// TIA Portal V19 export
// export: Created 2026-10-15T09:44:24.662474Z, ExportSetting WithDefaults, DisplayName Totally Integrated Automation Portal, DisplayVersion V19, DisplayName TIA Portal Openness, DisplayVersion V19, DisplayName TIA Portal Version Control Interface, DisplayVersion V19, DisplayName STEP 7 Professional, DisplayVersion V19, DisplayName STEP 7 Safety, DisplayVersion V19, DisplayName WinCC Basic/Comfort/Advanced, DisplayVersion V19, DisplayName WinCC Unified, DisplayVersion V19
FUNCTION "ROLL_PB20" : Void   // FC28, SCL
{ S7_Optimized_Access := 'TRUE' }
VERSION : 0.1
// stored: AutoNumber true, IsIECCheckEnabled false, SetENOAutomatically false, UDAEnableTagReadback false
   VAR_TEMP
      r : Bool;
      a1 : Word;
      a2 : Word;
      activeDataBlock : Int;
      comparisonResults : Array[0..0] of Bool;
   END_VAR
BEGIN

   #r := FALSE;
   #a1 := W#16#0000;
   #a2 := W#16#0000;
   #activeDataBlock := 0;
   // PB20, STEP 5 network 1
   #activeDataBlock := 15;
   // PB20, STEP 5 network 2
   #r := ((NOT "ROLL_IO".Input[7, 0]) AND (("ROLL_IO".Input[0, 1] AND "ROLL_State".M[190, 6] AND "ROLL_State".M[26, 5] AND "ROLL_State".M[4, 1]) OR ("ROLL_IO".Input[0, 2] AND "ROLL_State".M[0, 3])) AND "ROLL_State".M[4, 1]);
   "ROLL_State".M[8, 0] := #r;
   // PB20, STEP 5 network 3
   #r := ((NOT "ROLL_IO".Input[7, 1]) AND "ROLL_IO".Input[0, 2] AND "ROLL_IO".Input[1, 6] AND "ROLL_State".M[4, 1] AND "ROLL_State".S5Timers[61].Q);
   IF #r THEN
       "ROLL_State".M[8, 1] := TRUE;
   END_IF;
   #r := "ROLL_State".M[3, 1];
   IF #r THEN
       "ROLL_State".M[8, 1] := FALSE;
   END_IF;
   // PB20, STEP 5 network 4
   #a2 := #a1;
   #a1 := "ROLL_GetDW"(DbNumber := #activeDataBlock, Index := 61);
   #r := ((NOT "ROLL_IO".Input[7, 1]) AND "ROLL_IO".Input[0, 2] AND "ROLL_IO".Input[3, 1]);
   "ROLL_TimerOp"(Number := 61,
                  Operation := 0,
                  Signal := #r,
                  Preset := #a1);
   #r := ("ROLL_State".M[3, 1] AND "ROLL_State".M[4, 1]);
   "ROLL_TimerOp"(Number := 61,
                  Operation := 2,
                  Signal := #r,
                  Preset := #a1);
   // PB20, STEP 5 network 5
   #r := ((NOT "ROLL_IO".Input[7, 2]) AND "ROLL_State".S5Timers[55].Q);
   IF #r THEN
       "ROLL_State".M[8, 2] := TRUE;
   END_IF;
   #r := "ROLL_State".M[3, 1];
   IF #r THEN
       "ROLL_State".M[8, 2] := FALSE;
   END_IF;
   // PB20, STEP 5 network 6
   #a2 := #a1;
   #a1 := "ROLL_GetDW"(DbNumber := #activeDataBlock, Index := 55);
   #r := ((NOT "ROLL_IO".Input[7, 2]) AND (NOT "ROLL_State".M[8, 2]) AND "ROLL_State".M[4, 1]);
   "ROLL_TimerOp"(Number := 55,
                  Operation := 0,
                  Signal := #r,
                  Preset := #a1);
   // PB20, STEP 5 network 7
   #r := ((NOT "ROLL_IO".Input[7, 3]) AND "ROLL_IO".Output[21, 6] AND "ROLL_State".S5Timers[60].Q);
   IF #r THEN
       "ROLL_State".M[8, 3] := TRUE;
   END_IF;
   #r := "ROLL_State".M[3, 1];
   IF #r THEN
       "ROLL_State".M[8, 3] := FALSE;
   END_IF;
   // PB20, STEP 5 network 8
   #a2 := #a1;
   #a1 := "ROLL_GetDW"(DbNumber := #activeDataBlock, Index := 60);
   #r := ((NOT "ROLL_IO".Input[7, 3]) AND "ROLL_IO".Output[21, 6] AND "ROLL_IO".Input[3, 1]);
   "ROLL_TimerOp"(Number := 60,
                  Operation := 0,
                  Signal := #r,
                  Preset := #a1);
   // PB20, STEP 5 network 9
   #a2 := #a1;
   #a1 := W#16#2010;
   #r := (NOT "ROLL_IO".Input[7, 4]);
   "ROLL_TimerOp"(Number := 88,
                  Operation := 0,
                  Signal := #r,
                  Preset := #a1);
   // PB20, STEP 5 network 10
   #r := ((NOT "ROLL_IO".Input[7, 4]) AND "ROLL_State".M[4, 1] AND "ROLL_State".S5Timers[88].Q);
   "ROLL_State".M[8, 4] := #r;
   // PB20, STEP 5 network 11
   #r := (("ROLL_State".M[25, 0] OR "ROLL_State".M[25, 1]) AND "ROLL_IO".Input[0, 1] AND "ROLL_State".M[190, 6] AND "ROLL_State".M[4, 1] AND "ROLL_State".S5Timers[96].Q);
   IF #r THEN
       "ROLL_State".M[8, 5] := TRUE;
   END_IF;
   #r := "ROLL_State".M[3, 1];
   IF #r THEN
       "ROLL_State".M[8, 5] := FALSE;
   END_IF;
   // PB20, STEP 5 network 12
   #r := ((NOT "ROLL_IO".Input[9, 0]) AND ("ROLL_IO".Input[1, 6] OR "ROLL_IO".Input[1, 7]) AND "ROLL_IO".Input[9, 6]);
   IF #r THEN
       "ROLL_State".M[12, 4] := TRUE;
   END_IF;
   #r := "ROLL_State".M[3, 1];
   IF #r THEN
       "ROLL_State".M[12, 4] := FALSE;
   END_IF;
   // PB20, STEP 5 network 13
   #r := ((NOT "ROLL_IO".Input[9, 3]) AND ("ROLL_IO".Input[1, 6] OR "ROLL_IO".Input[1, 7]) AND "ROLL_IO".Input[9, 6]);
   IF #r THEN
       "ROLL_State".M[12, 5] := TRUE;
   END_IF;
   #r := "ROLL_State".M[3, 1];
   IF #r THEN
       "ROLL_State".M[12, 5] := FALSE;
   END_IF;
   // PB20, STEP 5 network 14
   #r := ((NOT "ROLL_IO".Input[9, 7]) AND ("ROLL_IO".Input[1, 6] OR "ROLL_IO".Input[1, 7]));
   IF #r THEN
       "ROLL_State".M[12, 6] := TRUE;
   END_IF;
   #r := "ROLL_State".M[3, 1];
   IF #r THEN
       "ROLL_State".M[12, 6] := FALSE;
   END_IF;
   // PB20, STEP 5 network 15
   #r := (NOT "ROLL_IO".Input[9, 6]);
   IF #r THEN
       "ROLL_State".M[12, 7] := TRUE;
   END_IF;
   #r := ("ROLL_IO".Input[9, 6] AND "ROLL_State".M[3, 1]);
   IF #r THEN
       "ROLL_State".M[12, 7] := FALSE;
   END_IF;
   // PB20, STEP 5 network 16
   #a2 := #a1;
   #a1 := "ROLL_GetDW"(DbNumber := #activeDataBlock, Index := 56);
   #r := (NOT "ROLL_IO".Input[7, 1]);
   "ROLL_TimerOp"(Number := 56,
                  Operation := 1,
                  Signal := #r,
                  Preset := #a1);
   // PB20, STEP 5 network 17
   #a2 := #a1;
   #a1 := "ROLL_GetDW"(DbNumber := #activeDataBlock, Index := 65);
   #r := (NOT "ROLL_IO".Input[7, 3]);
   "ROLL_TimerOp"(Number := 65,
                  Operation := 0,
                  Signal := #r,
                  Preset := #a1);
   // PB20, STEP 5 network 18
   #a2 := #a1;
   #a1 := W#16#2020;
   #r := "ROLL_IO".Input[7, 3];
   "ROLL_TimerOp"(Number := 66,
                  Operation := 1,
                  Signal := #r,
                  Preset := #a1);
   // PB20, STEP 5 network 19
   #a2 := #a1;
   #a1 := "ROLL_GetDW"(DbNumber := #activeDataBlock, Index := 67);
   #r := ("ROLL_IO".Input[7, 3] AND "ROLL_State".M[150, 1]);
   "ROLL_TimerOp"(Number := 67,
                  Operation := 0,
                  Signal := #r,
                  Preset := #a1);
   // PB20, STEP 5 network 20
   #a2 := #a1;
   #a1 := W#16#2005;
   #r := (NOT "ROLL_IO".Input[7, 5]);
   "ROLL_TimerOp"(Number := 96,
                  Operation := 0,
                  Signal := #r,
                  Preset := #a1);
   // PB20, STEP 5 network 21
   #a2 := #a1;
   #a1 := W#16#2030;
   #r := "ROLL_IO".Input[7, 5];
   "ROLL_TimerOp"(Number := 97,
                  Operation := 0,
                  Signal := #r,
                  Preset := #a1);
   // PB20, STEP 5 network 22
   #r := (((NOT "ROLL_IO".Output[18, 5]) AND "ROLL_IO".Output[18, 4]) OR ((NOT "ROLL_IO".Output[18, 7]) AND "ROLL_IO".Output[18, 6]));
   "ROLL_State".M[149, 6] := #r;
   // PB20, STEP 5 network 23
   #a2 := #a1;
   #a1 := W#16#1010;
   #r := "ROLL_State".M[148, 4];
   "ROLL_TimerOp"(Number := 89,
                  Operation := 0,
                  Signal := #r,
                  Preset := #a1);
   // PB20, STEP 5 network 24
   #r := "ROLL_State".M[149, 6];
   IF #r THEN
       "ROLL_State".M[148, 4] := TRUE;
   END_IF;
   #r := "ROLL_State".S5Timers[89].Q;
   IF #r THEN
       "ROLL_State".M[148, 4] := FALSE;
   END_IF;
   // PB20, STEP 5 network 25
   #r := ("ROLL_IO".Input[8, 0] AND "ROLL_State".S5Timers[70].Q);
   "ROLL_State".M[147, 0] := #r;
   // PB20, STEP 5 network 26
   #a2 := #a1;
   #a1 := "ROLL_GetDW"(DbNumber := #activeDataBlock, Index := 75);
   #r := (NOT "ROLL_State".M[147, 0]);
   "ROLL_TimerOp"(Number := 75,
                  Operation := 0,
                  Signal := #r,
                  Preset := #a1);
   // PB20, STEP 5 network 27
   #r := "ROLL_State".M[0, 3];
   "ROLL_State".M[147, 1] := #r;
   // PB20, STEP 5 network 28
   #r := ("ROLL_IO".Input[8, 2] AND "ROLL_State".S5Timers[72].Q);
   "ROLL_State".M[147, 2] := #r;
   // PB20, STEP 5 network 29
   #a2 := #a1;
   #a1 := "ROLL_GetDW"(DbNumber := #activeDataBlock, Index := 77);
   #r := (NOT "ROLL_State".M[147, 2]);
   "ROLL_TimerOp"(Number := 77,
                  Operation := 0,
                  Signal := #r,
                  Preset := #a1);
   // PB20, STEP 5 network 30
   #r := "ROLL_State".M[0, 3];
   "ROLL_State".M[149, 0] := #r;
   // PB20, STEP 5 network 31
   #r := ("ROLL_State".M[147, 0] OR "ROLL_State".M[147, 2]);
   "ROLL_State".M[149, 1] := #r;
   // PB20, STEP 5 network 32
   #r := "ROLL_State".M[0, 3];
   "ROLL_State".M[149, 2] := #r;
   // PB20, STEP 5 network 33
   #r := ("ROLL_State".M[147, 0] AND "ROLL_State".M[147, 2]);
   "ROLL_State".M[149, 3] := #r;
   // PB20, STEP 5 network 34
   #r := ((NOT "ROLL_State".M[12, 6]) AND (NOT "ROLL_State".M[12, 7]) AND (NOT "ROLL_State".M[13, 4]) AND (NOT "ROLL_State".M[6, 0]) AND (NOT "ROLL_State".M[6, 2]) AND (NOT "ROLL_State".M[8, 2]) AND ("ROLL_IO".Input[1, 6] OR "ROLL_IO".Input[1, 7]) AND "ROLL_IO".Input[3, 1] AND "ROLL_IO".Input[7, 4] AND "ROLL_IO".Input[9, 6] AND "ROLL_IO".Input[9, 7] AND "ROLL_State".S5Timers[66].Q);
   "ROLL_State".M[150, 2] := #r;
   // PB20, STEP 5 network 35
   #r := ((NOT "ROLL_IO".Input[9, 2]) AND (NOT "ROLL_State".M[12, 4]) AND ("ROLL_IO".Output[18, 4] OR "ROLL_IO".Input[9, 1]) AND ("ROLL_State".M[149, 0] OR "ROLL_State".M[149, 1] OR "ROLL_State".M[149, 2] OR "ROLL_State".M[149, 3]) AND "ROLL_IO".Input[9, 0] AND "ROLL_State".M[150, 2]);
   "ROLL_IO".Output[18, 4] := #r;
   // PB20, STEP 5 network 36
   #r := ((NOT "ROLL_IO".Input[9, 2]) AND (NOT "ROLL_State".M[12, 4]) AND ("ROLL_IO".Output[18, 4] OR "ROLL_IO".Output[18, 5] OR "ROLL_IO".Input[9, 1]) AND ("ROLL_State".M[149, 2] OR "ROLL_State".M[149, 3]) AND "ROLL_IO".Input[9, 0] AND "ROLL_State".M[150, 2]);
   "ROLL_IO".Output[18, 5] := #r;
   // PB20, STEP 5 network 37
   #r := ((NOT "ROLL_IO".Input[9, 5]) AND (NOT "ROLL_State".M[12, 5]) AND ("ROLL_IO".Output[18, 6] OR "ROLL_IO".Input[9, 4]) AND ("ROLL_State".M[149, 1] OR "ROLL_State".M[149, 2] OR "ROLL_State".M[149, 3]) AND "ROLL_IO".Input[9, 3] AND "ROLL_State".M[150, 2]);
   "ROLL_IO".Output[18, 6] := #r;
   // PB20, STEP 5 network 38
   #r := ((NOT "ROLL_IO".Input[9, 5]) AND (NOT "ROLL_State".M[12, 5]) AND ("ROLL_IO".Output[18, 6] OR "ROLL_IO".Output[18, 7] OR "ROLL_IO".Input[9, 4]) AND "ROLL_IO".Input[9, 3] AND "ROLL_State".M[149, 3] AND "ROLL_State".M[150, 2]);
   "ROLL_IO".Output[18, 7] := #r;
   // PB20, STEP 5 network 39
   #r := ((NOT "ROLL_State".M[147, 0]) AND "ROLL_State".M[147, 2] AND "ROLL_State".S5Timers[75].Q);
   "ROLL_IO".Output[21, 0] := #r;
   // PB20, STEP 5 network 40
   #r := ((NOT "ROLL_State".M[147, 2]) AND "ROLL_State".M[147, 0] AND "ROLL_State".S5Timers[77].Q);
   "ROLL_IO".Output[21, 2] := #r;
   // PB20, STEP 5 network 41
   #r := "ROLL_State".M[190, 6];
   IF #r THEN
       "ROLL_State".M[150, 0] := TRUE;
   END_IF;
   #r := ((NOT "ROLL_IO".Input[0, 1]) OR (NOT "ROLL_IO".Input[7, 1]) OR (NOT "ROLL_IO".Input[7, 2]) OR (NOT "ROLL_State".M[27, 5]) OR "ROLL_IO".Input[7, 3] OR "ROLL_State".M[190, 5]);
   IF #r THEN
       "ROLL_State".M[150, 0] := FALSE;
   END_IF;
   // PB20, STEP 5 network 42
   #a2 := #a1;
   #a1 := W#16#2020;
   #r := "ROLL_IO".Input[7, 1];
   "ROLL_TimerOp"(Number := 57,
                  Operation := 1,
                  Signal := #r,
                  Preset := #a1);
   // PB20, STEP 5 network 43
   #r := ((NOT "ROLL_State".M[13, 4]) AND (NOT "ROLL_State".S5Timers[61].Q) AND (((NOT "ROLL_IO".Input[7, 3]) AND "ROLL_State".S5Timers[65].Q) OR ((NOT "ROLL_State".S5Timers[67].Q) AND "ROLL_State".M[150, 1])) AND "ROLL_IO".Input[0, 2] AND "ROLL_IO".Input[3, 1] AND "ROLL_IO".Input[7, 2] AND "ROLL_State".S5Timers[57].Q);
   "ROLL_State".M[150, 1] := #r;
   // PB20, STEP 5 network 44
   #r := ("ROLL_State".M[150, 0] OR "ROLL_State".M[150, 1]);
   "ROLL_IO".Output[21, 6] := #r;
   // PB20, STEP 5 network 45
   #r := ((((NOT "ROLL_IO".Input[7, 4]) AND "ROLL_IO".Input[7, 5]) OR ((NOT "ROLL_State".S5Timers[106].Q) AND "ROLL_State".M[148, 6]) OR (NOT "ROLL_IO".Input[7, 1])) AND "ROLL_IO".Input[0, 2] AND "ROLL_IO".Input[1, 6] AND "ROLL_IO".Input[7, 0]);
   "ROLL_State".M[148, 6] := #r;
   // PB20, STEP 5 network 46
   #r := (((NOT "ROLL_State".M[151, 0]) AND (NOT "ROLL_State".M[151, 1]) AND (NOT "ROLL_State".M[151, 2]) AND (NOT "ROLL_State".M[151, 3])) OR ((NOT "ROLL_State".M[152, 3]) AND "ROLL_State".M[151, 3] AND "ROLL_State".M[153, 3] AND "ROLL_State".S5Timers[105].Q));
   IF #r THEN
       "ROLL_State".M[151, 0] := TRUE;
   END_IF;
   #r := ("ROLL_State".M[151, 1] OR "ROLL_State".M[151, 2]);
   IF #r THEN
       "ROLL_State".M[151, 0] := FALSE;
   END_IF;
   // PB20, STEP 5 network 47
   #a2 := #a1;
   #a1 := "ROLL_GetDW"(DbNumber := #activeDataBlock, Index := 102);
   #r := "ROLL_State".M[151, 0];
   "ROLL_TimerOp"(Number := 102,
                  Operation := 0,
                  Signal := #r,
                  Preset := #a1);
   // PB20, STEP 5 network 48
   #r := ((NOT "ROLL_State".S5Timers[106].Q) AND "ROLL_State".M[151, 0]);
   IF #r THEN
       "ROLL_State".M[152, 0] := TRUE;
   END_IF;
   #r := ((NOT "ROLL_State".M[148, 6]) OR "ROLL_State".S5Timers[106].Q);
   IF #r THEN
       "ROLL_State".M[152, 0] := FALSE;
   END_IF;
   // PB20, STEP 5 network 49
   #r := ("ROLL_IO".Output[21, 5] AND "ROLL_State".M[152, 0]);
   IF #r THEN
       "ROLL_State".M[153, 0] := TRUE;
   END_IF;
   #r := (NOT "ROLL_State".M[151, 0]);
   IF #r THEN
       "ROLL_State".M[153, 0] := FALSE;
   END_IF;
   // PB20, STEP 5 network 50
   #r := ((NOT "ROLL_State".M[152, 0]) AND "ROLL_State".M[151, 0] AND "ROLL_State".M[153, 0] AND "ROLL_State".S5Timers[102].Q);
   IF #r THEN
       "ROLL_State".M[151, 1] := TRUE;
   END_IF;
   #r := "ROLL_State".M[151, 2];
   IF #r THEN
       "ROLL_State".M[151, 1] := FALSE;
   END_IF;
   // PB20, STEP 5 network 51
   #a2 := #a1;
   #a1 := "ROLL_GetDW"(DbNumber := #activeDataBlock, Index := 103);
   #r := "ROLL_State".M[151, 1];
   "ROLL_TimerOp"(Number := 103,
                  Operation := 0,
                  Signal := #r,
                  Preset := #a1);
   // PB20, STEP 5 network 52
   #r := ((NOT "ROLL_State".S5Timers[106].Q) AND "ROLL_State".M[151, 1]);
   IF #r THEN
       "ROLL_State".M[152, 1] := TRUE;
   END_IF;
   #r := ((NOT "ROLL_State".M[148, 6]) OR "ROLL_State".S5Timers[106].Q);
   IF #r THEN
       "ROLL_State".M[152, 1] := FALSE;
   END_IF;
   // PB20, STEP 5 network 53
   #r := ("ROLL_IO".Output[20, 6] AND "ROLL_State".M[152, 1]);
   IF #r THEN
       "ROLL_State".M[153, 1] := TRUE;
   END_IF;
   #r := (NOT "ROLL_State".M[151, 1]);
   IF #r THEN
       "ROLL_State".M[153, 1] := FALSE;
   END_IF;
   // PB20, STEP 5 network 54
   #r := ((NOT "ROLL_State".M[152, 1]) AND "ROLL_State".M[151, 1] AND "ROLL_State".M[153, 1] AND "ROLL_State".S5Timers[103].Q);
   IF #r THEN
       "ROLL_State".M[151, 2] := TRUE;
   END_IF;
   #r := "ROLL_State".M[151, 3];
   IF #r THEN
       "ROLL_State".M[151, 2] := FALSE;
   END_IF;
   // PB20, STEP 5 network 55
   #a2 := #a1;
   #a1 := W#16#0002;
   #r := "ROLL_State".M[151, 2];
   "ROLL_TimerOp"(Number := 104,
                  Operation := 0,
                  Signal := #r,
                  Preset := #a1);
   // PB20, STEP 5 network 56
   #r := ((NOT "ROLL_State".S5Timers[106].Q) AND "ROLL_State".M[151, 2]);
   IF #r THEN
       "ROLL_State".M[152, 2] := TRUE;
   END_IF;
   #r := ((NOT "ROLL_State".M[148, 6]) OR "ROLL_State".S5Timers[106].Q);
   IF #r THEN
       "ROLL_State".M[152, 2] := FALSE;
   END_IF;
   // PB20, STEP 5 network 57
   #r := ("ROLL_State".M[0, 4] AND "ROLL_State".M[152, 2]);
   IF #r THEN
       "ROLL_State".M[153, 2] := TRUE;
   END_IF;
   #r := (NOT "ROLL_State".M[151, 2]);
   IF #r THEN
       "ROLL_State".M[153, 2] := FALSE;
   END_IF;
   // PB20, STEP 5 network 58
   #r := ((NOT "ROLL_State".M[152, 2]) AND "ROLL_State".M[151, 2] AND "ROLL_State".M[153, 2] AND "ROLL_State".S5Timers[104].Q);
   IF #r THEN
       "ROLL_State".M[151, 3] := TRUE;
   END_IF;
   #r := "ROLL_State".M[151, 0];
   IF #r THEN
       "ROLL_State".M[151, 3] := FALSE;
   END_IF;
   // PB20, STEP 5 network 59
   #a2 := #a1;
   #a1 := W#16#0002;
   #r := "ROLL_State".M[151, 3];
   "ROLL_TimerOp"(Number := 105,
                  Operation := 0,
                  Signal := #r,
                  Preset := #a1);
   // PB20, STEP 5 network 60
   #r := ((NOT "ROLL_State".S5Timers[106].Q) AND "ROLL_State".M[151, 3]);
   IF #r THEN
       "ROLL_State".M[152, 3] := TRUE;
   END_IF;
   #r := ((NOT "ROLL_State".M[148, 6]) OR "ROLL_State".S5Timers[106].Q);
   IF #r THEN
       "ROLL_State".M[152, 3] := FALSE;
   END_IF;
   // PB20, STEP 5 network 61
   #r := ("ROLL_State".M[0, 4] AND "ROLL_State".M[152, 3]);
   IF #r THEN
       "ROLL_State".M[153, 3] := TRUE;
   END_IF;
   #r := (NOT "ROLL_State".M[151, 3]);
   IF #r THEN
       "ROLL_State".M[153, 3] := FALSE;
   END_IF;
   // PB20, STEP 5 network 62
   #a2 := #a1;
   #a1 := W#16#2010;
   #r := ("ROLL_State".M[152, 0] OR "ROLL_State".M[152, 1] OR "ROLL_State".M[152, 2] OR "ROLL_State".M[152, 3]);
   "ROLL_TimerOp"(Number := 106,
                  Operation := 0,
                  Signal := #r,
                  Preset := #a1);
   // PB20, STEP 5 network 63
   #r := ((NOT "ROLL_IO".Output[21, 4]) AND "ROLL_IO".Output[19, 5] AND "ROLL_State".M[152, 0]);
   "ROLL_IO".Output[21, 5] := #r;
   // PB20, STEP 5 network 64
   #r := "ROLL_State".M[152, 1];
   "ROLL_State".M[240, 0] := #r;
   // PB20, STEP 5 network 65
   #r := ((NOT "ROLL_IO".Output[21, 5]) AND "ROLL_State".M[152, 2]);
   "ROLL_State".M[240, 0] := #r;
   // PB20, STEP 5 network 66
   #r := "ROLL_State".M[152, 3];
   "ROLL_State".M[240, 0] := #r;
   // PB20, STEP 5 network 67
   #a2 := #a1;
   #a1 := "ROLL_GetDW"(DbNumber := #activeDataBlock, Index := 107);
   #r := ("ROLL_IO".Output[21, 6] AND "ROLL_IO".Input[0, 2]);
   "ROLL_TimerOp"(Number := 107,
                  Operation := 1,
                  Signal := #r,
                  Preset := #a1);
   // PB20, STEP 5 network 68
   #r := ((("ROLL_IO".Output[21, 6] OR "ROLL_State".S5Timers[107].Q) AND "ROLL_IO".Input[0, 2]) OR ("ROLL_IO".Input[0, 1] AND "ROLL_State".M[190, 6] AND "ROLL_State".M[26, 6]));
   "ROLL_IO".Output[20, 5] := #r;
   // PB20, STEP 5 network 69
   RETURN;
END_FUNCTION
